ABB RobotStudio station: RS4.rsstn

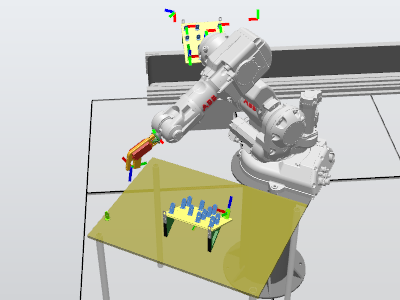
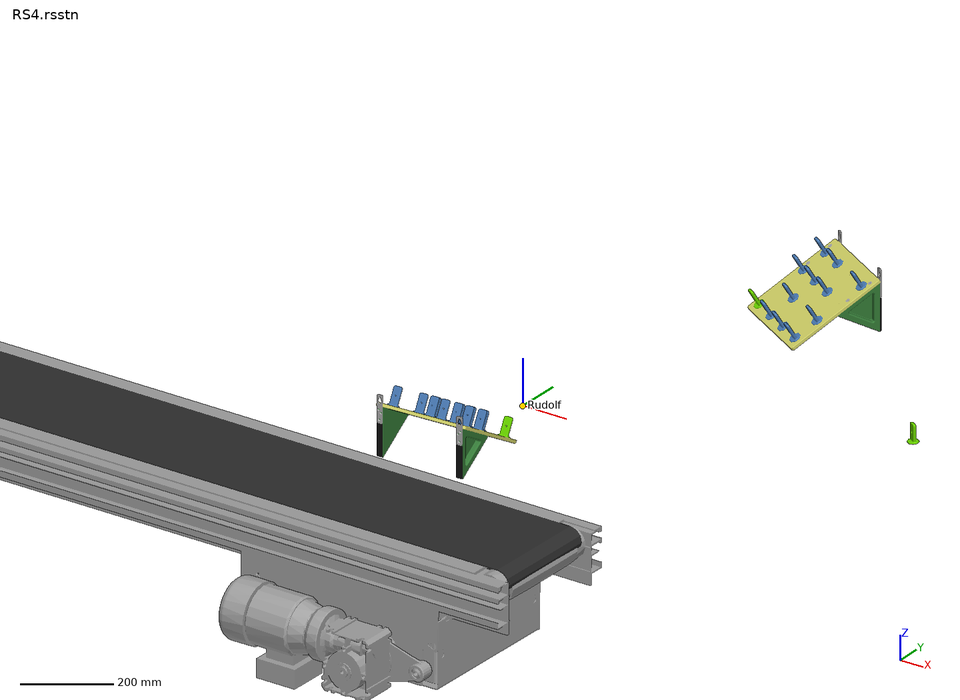
[picture v1: parts stored in the station drawn from their meshes, with robot base, taught points and paths (robot models come from the ABB library and are not in the file)]
Station RS4_tatem (saved by RobotStudio 25.5.11605.0)
Controller Rudolf, task T_ROB1: task frame (RAPID world) sits at (10, 680, 720) mm, rotated rx 0 ry 0 rz -30 deg in the station
Controller Rudolf
  mechanical unit ROB_1: Rudolf, 6 joints, base frame (0, 0, 0) mm
Layout (positions relative to the parent item):
  - PedestalR [part, from Libraries\Pedestal.rslib] at (10, 680, 0) mm, rotated rx 0 ry 0 rz 150 deg
  - TableR [part, from Libraries\Desk.rslib] at (193.4, 1497.66, 0) mm, rotated rx 0 ry 0 rz -120 deg
  - Rudolf [mechanism, from Libraries\IRB140_6_81_C_G_03.rslib] at (10, 680, 720) mm, rotated rx 0 ry 0 rz -30 deg; joint values [1.0472, 0.5236, 0, 0, -0.1745, 1.5708] (rad or m)
  - Spot welding tool UiS [part, from Libraries\Spot welding tool UiS.rslib] at (564.4, 1000.09, 1171.54) mm, rotated rx 110 ry 0 rz 120 deg
  - Board on table [part] at (358.49, 1103.75, 828) mm, rotated rx 0 ry 0 rz 60 deg, size 218.4 x 225 x 147.8 mm
  - Board on belt [part] at (278.92, 104.3, 964) mm, rotated rx 0 ry 0 rz -87 deg, size 218.4 x 225 x 147.8 mm
  - Conveyor [part] at (-998.97, -64.27, 804) mm, rotated rx 90 ry -1 rz -90 deg, size 568.5 x 300.9 x 1730 mm
  - FreePeg [part] at (800, 1000, 751) mm, rotated rx 0 ry 0 rz -30 deg, size 25 x 25 x 44 mm
Attachment: TableR is attached to PedestalR
Attachment: Spot welding tool UiS is attached to Rudolf / Link6
Attachment: wobjTestBoard is attached to Board on table
Attachment: wobjTestBoardOnBelt is attached to Board on belt
Station signals: DI doClose, DI doOpen
Station logic (signal -> signal, property => property):
  Norbert.doOpen -> SC_Gripper.diOpen
  Norbert.doClose -> SC_Gripper.diClose
  SC_Gripper.doClosed -> Norbert.diClosed
Targets, tools, work objects and paths stored in the station, written as RAPID:
! task T_ROB1
MODULE MainModule
  CONST speeddata v_SuperSlow:=[100,500,5000,1000];
  CONST speeddata v_fullpinne:=[5000,5000,5000,1000];
  CONST speeddata v_VeryFast:=[5000,5000,5000,1000];
  CONST speeddata v_VerySlow:=[ 100,500,5000,1000];
  VAR NUM tWait:=0.59;
  VAR speeddata speed_1:=[ 500,500,5000,1000];
  CONST speeddata v_Fast:=[1000,500,5000,1000];
  CONST speeddata v_Slow:=[ 200,500,5000,1000];
  PERS tooldata TatemTool1:=[TRUE,[[0,-48.3,153.5],[0,0,-0.5,0.866025404]],[0.3,[0,0,1],[1,0,0,0],0,0,0]];
  TASK PERS wobjdata wobjTestBoardOnBelt:=[FALSE,TRUE,"",[[599.763,-318.75,282.622],[0.265084,0.0713605,-0.252646,-0.927797]],[[0,0,0],[1,0,0,0]]];
  TASK PERS wobjdata wobjTableR:=[FALSE,TRUE,"",[[150,500,8],[1,0,0,0]],[[0,0,0],[1,0,0,0]]];
  CONST robtarget AboveTestBoard:=[[90,90,100],[0,1,0,0],[1,0,-1,1],[9E+09,9E+09,9E+09,9E+09,9E+09,9E+09]];
  CONST robtarget Peg_00:=[[0,0,0],[0,1,0,0],[1,0,-1,1],[9E+09,9E+09,9E+09,9E+09,9E+09,9E+09]];
  CONST robtarget Peg_03:=[[0,180,0],[0,1,0,0],[1,0,-1,1],[9E+09,9E+09,9E+09,9E+09,9E+09,9E+09]];
  CONST robtarget Peg_30:=[[180,0,0],[0,1,0,0],[0,-1,0,1],[9E+09,9E+09,9E+09,9E+09,9E+09,9E+09]];
  CONST robtarget Peg_33:=[[180,180,0],[0,1,0,0],[0,-1,0,1],[9E+09,9E+09,9E+09,9E+09,9E+09,9E+09]];
  TASK PERS wobjdata wobjTestBoard:=[FALSE,TRUE,"",[[599.763,-318.75,282.622],[0.265084,0.0713605,-0.252646,-0.927797]],[[0,0,0],[1,0,0,0]]];
  CONST jointtarget jCalibPos0:=[[0,0,0,0,0,0],[9E+09,9E+09,9E+09,9E+09,9E+09,9E+09]];
  CONST jointtarget jCalibPosR:=[[-60,30,0,0,-10,90],[9E+09,9E+09,9E+09,9E+09,9E+09,9E+09]];
  CONST jointtarget jCalibPosL:=[[60,30,0,0,-10,90],[9E+09,9E+09,9E+09,9E+09,9E+09,9E+09]];
  CONST speeddata vFast:=[1000,500,5000,1000];
  TASK PERS wobjdata wobjTestBoardOnTable:=[FALSE,TRUE,"",[[0,544,146],[0.965928085,0.258810616,0,0]],[[0,0,0],[1,0,0,0]]];
  CONST speeddata vSlow:=[ 200,500,5000,1000];
  VAR jointtarget jCalibPos:=[[0,0,0,0,0,0],[9E+09,9E+09,9E+09,9E+09,9E+09,9E+09]];
  PROC main()
    testPeg00;
    test4corners;
    WaitTime 0.1;
    MoveAbsJ jCalibPos0,v1000,z10,tool0;
  ENDPROC
  PROC initTatemTool()
  ENDPROC
  PROC test4corners()
    MoveAbsJ jCalibPos,vFast,z10,tool0;
    initTatemTool;
    MoveAbsJ jCalibPos,vFast,z10,tool0;
  ENDPROC
  PROC testPeg00()
    MoveAbsJ jCalibPos,vFast,z10,tool0;
    initTatemTool;
    MoveAbsJ jCalibPos,vFast,z10,tool0;
  ENDPROC
ENDMODULE

! task T_ROB1
MODULE trigtest
  CONST speeddata v_ToolSpeed:=[  50,500,5000,1000];
ENDMODULE

! task T_ROB1
MODULE LINKEDM
  PROC Linked_m()
  ENDPROC
ENDMODULE

